Staubli VAL3: utCommon.dtx

public bool bDisabled
public string sValue
public string sID
public string sOption{}
public string sItem
public string sPage
